FUNCTION_BLOCK RP (* Basic Function Block Type *)
  (* Standard: 61499-2 *)
  (* Version 0.0, 1/4/2020, prana, nxtControl GmbH, Template *)
  PACKAGE Main;
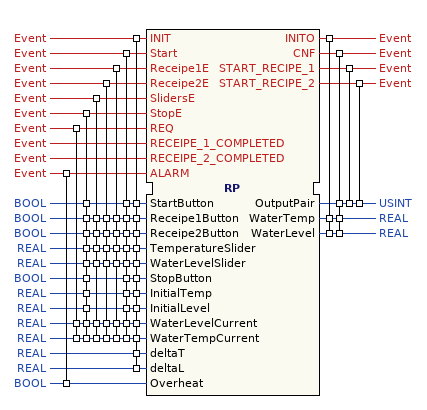
  EVENT_INPUT
    INIT WITH StartButton, Receipe1Button, Receipe2Button, TemperatureSlider, WaterLevelSlider, StopButton, InitialTemp, InitialLevel, WaterLevelCurrent, WaterTempCurrent, deltaT, deltaL;
    Start WITH StartButton, Receipe1Button, Receipe2Button, TemperatureSlider, WaterLevelSlider, StopButton, InitialTemp, InitialLevel, WaterLevelCurrent, WaterTempCurrent;
    Receipe1E WITH Receipe1Button, Receipe2Button, TemperatureSlider, WaterLevelSlider, WaterLevelCurrent, WaterTempCurrent; (* Initialization Request *)
    Receipe2E WITH Receipe1Button, Receipe2Button, TemperatureSlider, WaterLevelSlider, WaterLevelCurrent, WaterTempCurrent; (* Normal Execution Request *)
    SlidersE WITH Receipe1Button, Receipe2Button, TemperatureSlider, WaterLevelSlider, WaterLevelCurrent, WaterTempCurrent;
    StopE WITH StartButton, Receipe1Button, Receipe2Button, TemperatureSlider, WaterLevelSlider, StopButton, InitialTemp, InitialLevel, WaterLevelCurrent, WaterTempCurrent;
    REQ WITH WaterLevelCurrent, WaterTempCurrent;
    RECEIPE_1_COMPLETED;
    RECEIPE_2_COMPLETED;
    ALARM WITH Overheat;
  END_EVENT
  EVENT_OUTPUT
    INITO WITH WaterLevel, WaterTemp; (* Initialization Confirm *)
    CNF WITH WaterTemp, WaterLevel, OutputPair; (* Execution Confirmation *)
    START_RECIPE_1 WITH OutputPair;
    START_RECIPE_2 WITH OutputPair;
  END_EVENT
  VAR_INPUT
    StartButton : BOOL;
    Receipe1Button : BOOL; (* Input event qualifier *)
    Receipe2Button : BOOL;
    TemperatureSlider : REAL;
    WaterLevelSlider : REAL;
    StopButton : BOOL;
    InitialTemp : REAL;
    InitialLevel : REAL;
    WaterLevelCurrent : REAL;
    WaterTempCurrent : REAL;
    deltaT : REAL;
    deltaL : REAL;
    Overheat : BOOL;
  END_VAR
  VAR_OUTPUT
    OutputPair : USINT := 2;
    WaterTemp : REAL;
    WaterLevel : REAL; (* Output event qualifier *)
  END_VAR
  VAR
    X1 : REAL := 165.50;
    Y1 : REAL := 50.00;
    X2 : REAL := 250.50;
    Y2 : REAL := 68.96;
  END_VAR
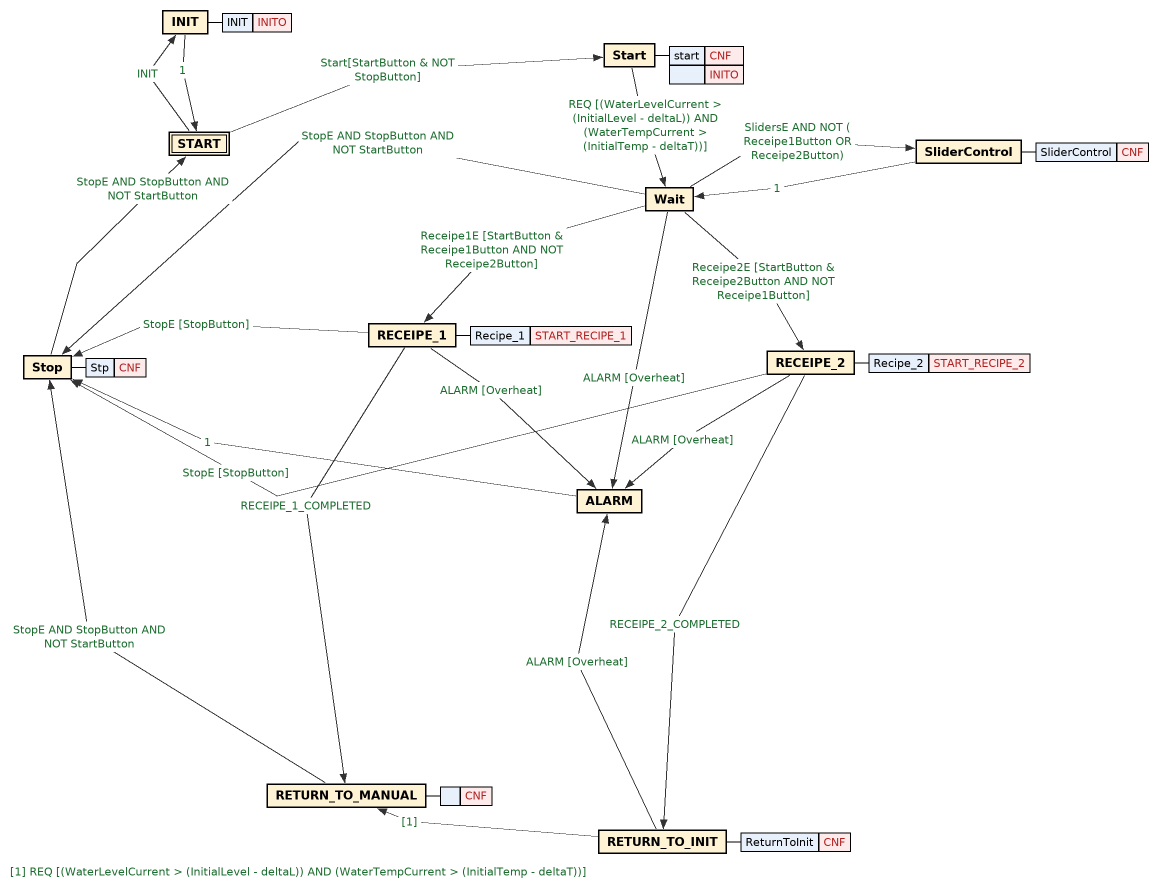
  EC_STATES
    START; (* Initial State *)
    SliderControl : SliderControl -> CNF;
    Start : start -> CNF, -> INITO;
    Stop : Stp -> CNF;
    INIT : INIT -> INITO;
    RECEIPE_1 : Recipe_1 -> START_RECIPE_1;
    RETURN_TO_MANUAL : -> CNF;
    RECEIPE_2 : Recipe_2 -> START_RECIPE_2;
    Wait;
    RETURN_TO_INIT : ReturnToInit -> CNF;
    ALARM;
  END_STATES
  EC_TRANSITIONS
    Wait TO SliderControl := SlidersE AND NOT ( Receipe1Button OR Receipe2Button);
    START TO Start := Start[StartButton & NOT StopButton];
    Wait TO RECEIPE_1 := Receipe1E [StartButton & Receipe1Button AND NOT Receipe2Button];
    Stop TO START := StopE AND StopButton AND NOT StartButton;
    START TO INIT := INIT;
    INIT TO START := 1;
    RECEIPE_1 TO RETURN_TO_MANUAL := RECEIPE_1_COMPLETED;
    RECEIPE_2 TO RETURN_TO_INIT := RECEIPE_2_COMPLETED;
    Wait TO RECEIPE_2 := Receipe2E [StartButton & Receipe2Button AND NOT Receipe1Button];
    RETURN_TO_MANUAL TO Stop := StopE AND StopButton AND NOT StartButton;
    SliderControl TO Wait := 1;
    Start TO Wait := REQ [(WaterLevelCurrent > (InitialLevel - deltaL)) AND (WaterTempCurrent > (InitialTemp - deltaT))];
    Wait TO Stop := StopE AND StopButton AND NOT StartButton;
    RETURN_TO_INIT TO RETURN_TO_MANUAL := REQ [(WaterLevelCurrent > (InitialLevel - deltaL)) AND (WaterTempCurrent > (InitialTemp - deltaT))];
    RECEIPE_1 TO Stop := StopE [StopButton];
    RECEIPE_1 TO ALARM := ALARM [Overheat];
    RECEIPE_2 TO ALARM := ALARM [Overheat];
    RETURN_TO_INIT TO ALARM := ALARM [Overheat];
    ALARM TO Stop := 1;
    RECEIPE_2 TO Stop := StopE [StopButton];
    Wait TO ALARM := ALARM [Overheat];
  END_TRANSITIONS
  ALGORITHM INIT IN ST: (* Initialization algorithm *)
;
OutputPair := 2;
  END_ALGORITHM
  ALGORITHM SliderControl IN ST:
WaterLevel := WaterLevelSlider;
WaterTemp := TemperatureSlider;
  END_ALGORITHM
  ALGORITHM start IN ST:
WaterLevel := InitialLevel;
WaterTemp := InitialTemp;
OutputPair := 2;
  END_ALGORITHM
  ALGORITHM Stp IN ST:
WaterLevel := 0;
WaterTemp := 0;
OutputPair := 2;
  END_ALGORITHM
  ALGORITHM X1 IN ST:
WaterLevel := X1;
WaterTemp := Y2;
  END_ALGORITHM
  ALGORITHM X2 IN ST:
WaterLevel := X2;
WaterTemp := Y2;
  END_ALGORITHM
  ALGORITHM Drain IN ST:
WaterLevel := 0;
WaterTemp := 0;
  END_ALGORITHM
  ALGORITHM Recipe_1 IN ST:
;
OutputPair := 0;
  END_ALGORITHM
  ALGORITHM ManualOutput IN ST:
;
OutputPair := 2;
  END_ALGORITHM
  ALGORITHM Recipe_2 IN ST:
;
OutputPair := 1;
  END_ALGORITHM
  ALGORITHM ReturnToInit IN ST:
;
WaterLevel := InitialLevel;
WaterTemp := InitialTemp;
OutputPair := 2;
  END_ALGORITHM
END_FUNCTION_BLOCK
